(* IEC 61131-3 sources: TetherPLC/tests/mixed, 3 files *)

(* ---- lib.st ---- *)
FUNCTION_BLOCK StFb
VAR_INPUT X : LREAL; END_VAR
VAR_OUTPUT Y : LREAL; END_VAR
Y := X * 2.0;
END_FUNCTION_BLOCK

FUNCTION StFn : LREAL
VAR_INPUT A : LREAL; END_VAR
StFn := A + 10.0;
END_FUNCTION

(* ---- dup.st ---- *)
PROGRAM Main
VAR x : BOOL; END_VAR
x := TRUE;
END_PROGRAM

(* ---- stprog.st ---- *)
PROGRAM StProg
VAR f : FbdFb; r : BOOL; END_VAR
f(IN := FALSE);
r := f.OUT;
END_PROGRAM
